TYPE ST_EL28x9 :
STRUCT
	//16CH DO, PNP 24VDC/0.5A  - 2809
	//16CH DO, GND-SW, 24VDC/0.5A - 2889
	
	State	AT %I*: UINT;

	q_ch1	AT %Q*: BOOL;
	q_ch2	AT %Q*: BOOL;
	q_ch3	AT %Q*: BOOL;
	q_ch4	AT %Q*: BOOL;
	q_ch5	AT %Q*: BOOL;
	q_ch6	AT %Q*: BOOL;
	q_ch7	AT %Q*: BOOL;
	q_ch8	AT %Q*: BOOL;
	
	q_ch9	AT %Q*: BOOL;
	q_ch10	AT %Q*: BOOL;
	q_ch11	AT %Q*: BOOL;
	q_ch12	AT %Q*: BOOL;
	q_ch13	AT %Q*: BOOL;
	q_ch14	AT %Q*: BOOL;
	q_ch15	AT %Q*: BOOL;
	q_ch16	AT %Q*: BOOL;
	
(*	
	bit_ch1	AT %Q*: BIT;
	bit_ch2	AT %Q*: BIT;
	bit_ch3	AT %Q*: BIT;
	bit_ch4	AT %Q*: BIT;
	bit_ch5	AT %Q*: BIT;
	bit_ch6	AT %Q*: BIT;
	bit_ch7	AT %Q*: BIT;
	bit_ch8	AT %Q*: BIT;
	
	bit_ch9		AT %Q*: BIT;
	bit_ch10	AT %Q*: BIT;
	bit_ch11	AT %Q*: BIT;
	bit_ch12	AT %Q*: BIT;
	bit_ch13	AT %Q*: BIT;
	bit_ch14	AT %Q*: BIT;
	bit_ch15	AT %Q*: BIT;
	bit_ch16	AT %Q*: BIT;
*)	
	
	
	
END_STRUCT
END_TYPE

(* stored: Version 1.1.0.1, ProductVersion 3.1.4024.12
   DUT ST_EL28x9: Id {61437754-2ae3-4153-9773-2ea41f9c1c3c} *)
